(* IEC 61131-3 sources: Lasal-MCP/examples/SampleSource/LASALScreenAdvancedSolution/LASALScreenAdvancedSolution/LASALScreenAdvacnedSolution/Stations/Terminal/HMI/Class/DataRecord, 1 file *)

(* ---- DataRecord.st ---- *)
(*!
<Class
	Name               = "DataRecord"
	Revision           = "0.0"
	RealtimeTask       = "false"
	CyclicTask         = "false"
	BackgroundTask     = "false"
	Sigmatek           = "false"
	OSInterface        = "false"
	HighPriority       = "false"
	Automatic          = "false"
	UpdateMode         = "Prescan"
	SharedCommandTable = "true"
	Objectsize         = "(450,360)">
	<Channels>
		<Server Name="CoordX" Visualized="true" Initialize="false" WriteProtected="true" Retentive="false"/>
		<Server Name="CoordY" Visualized="true" Initialize="false" WriteProtected="true" Retentive="false"/>
		<Server Name="IntError" Visualized="false" Initialize="false" WriteProtected="true" Retentive="false"/>
		<Client Name="_Grafix" Required="false" Internal="false"/>
		<Client Name="_StdLib" Required="false" Internal="false"/>
		<Client Name="AllocateSize" Required="false" Internal="false" DefValue="4 KB"/>
	</Channels>
	<Network Name="DataRecord">
		<!-- List of Components in this network -->
		<Components>
			<Object
				Name       = "_base"
				Class      = "_MyIO"
				Position   = "(218,120)"
				Visualized = "true"
				Remotely   = "true">
				<Channels>
					<Server Name="Refresh"/>
					<Server Name="Server0"/>
					<Client Name="Graphic"/>
					<Client Name="Lse"/>
				</Channels>
			</Object>
		</Components>
		<Comments>
		</Comments>
		<!-- List of Connections in this network -->
		<Connections>
			<Connection Source="this.Server0" Destination="_base.Server0" Vertices="(706,210),(534,210),"/>
			<Connection Source="this.Refresh" Destination="_base.Refresh" Vertices="(706,270),(534,270),"/>
			<Connection Source="_base.Lse" Destination="this.Lse" Vertices="(218,210),(38,210),"/>
		</Connections>
		<!-- Headerfiles -->
		<Options>
		</Options>
	</Network>
</Class>
*)
#pragma using _MyIO

DataRecord : CLASS
: _MyIO
  //Servers:
	CoordX 	: SvrCh_DINT;
	CoordY 	: SvrCh_DINT;
	IntError 	: SvrCh_DINT;
  //Clients:
	_Grafix 	: CltChCmd__Grafix;
	_StdLib 	: CltChCmd__StdLib;
	AllocateSize 	: CltCh_UDINT;
  //Variables:
		pStart 	: ^_DOT;
		pCheck 	: ^_DOT;
		pAct 	: ^_DOT;
		NoOfBufferEntries 	: UDINT;
		MaxNoOfBufferEntries 	: UDINT;
		Delete 	: DINT;
		pError 	: ^void;
  //Functions:

	FUNCTION VIRTUAL GLOBAL Init;
				//! <Function Comment="this method will be called once when the focus will be given to this object" Name="GetFocus"/>
	FUNCTION __CDECL VIRTUAL GLOBAL GetFocus
		VAR_INPUT
			pio 	: ^_IO;			//! <Variable Comment="pointer to _IO information" Name="GetFocus.pio"/>
		END_VAR
		VAR_OUTPUT
			retcode (EAX) 	: _DOIT;			//! <Variable Comment="return _IFAILED if you dont want to get the focus on the other hand _IDLE" Name="GetFocus.retcode"/>
		END_VAR;
				//! <Function Comment="this method is called everytime when the input is active and a event occured" Name="GetEvent"/>
	FUNCTION __CDECL VIRTUAL GLOBAL GetEvent
		VAR_INPUT
			ped 	: ^_EDITOR;			//! <Variable Comment="pointer to _EDITOR information" Name="GetEvent.ped"/>
			pe 	: ^_EVENT;			//! <Variable Comment="pointer to _EVENT information" Name="GetEvent.pe"/>
		END_VAR
		VAR_OUTPUT
			retcode (EAX) 	: _DOIT;			//! <Variable Comment="for the returnstatement there are 3 different possibilities&#13;&#10;  _IDLE ..... the system should goon like it is (system goes on)&#13;&#10;  _IDIDIT ... i did it (system is ready)&#13;&#10;  _IFAILED .. i tried to do my best, but i failed (system is ready)&#13;&#10;" Name="GetEvent.retcode"/>
		END_VAR;
				//! <Function Comment="this method is called everytime when system wants to redraw the io" Name="Draw"/>
	FUNCTION __CDECL VIRTUAL GLOBAL Draw
		VAR_INPUT
			pio 	: ^_IO;			//! <Variable Comment="pointer to _IO information" Name="Draw.pio"/>
			pr 	: ^_RESULT;			//! <Variable Comment="pointer to _RESULT information" Name="Draw.pr"/>
			pv 	: ^_VARIABLE;			//! <Variable Comment="pointer to io _VARIABLE information" Name="Draw.pv"/>
			input 	: BOOL;			//! <Variable Comment="TRUE it&apos;s an input&#13;&#10;FALSE it&apos;s an output" Name="Draw.input"/>
		END_VAR
		VAR_OUTPUT
			retcode (EAX) 	: _DOIT;			//! <Variable Comment="for the returnstatement there are 3 different possibilities&#13;&#10;  _IDLE ..... the system should goon like it is (system goes on)&#13;&#10;  _IDIDIT ... i did it (system is ready)&#13;&#10;  _IFAILED .. i tried to do my best, but i failed (system is re" Name="Draw.retcode"/>
		END_VAR;
				//! <Function Comment="this method is called everytime when system wants to get data for defined io.&#13;&#10;&#13;&#10;pr ........ &#13;&#10;pio ....... pointer to io information&#13;&#10;pv ........ pointer to io variableinformation&#13;&#10;input ..... TRUE it&apos;s an input / FALSE it&apos;s an output&#13;&#10;&#13;&#10;for the returnstatement there are 3 different possibilities&#13;&#10;_IDLE ..... the system should goon like it is (system goes on)&#13;&#10;_IDIDIT ... i did it (system is ready)&#13;&#10;_IFAILED .. i tried to do my best, but i failed (system is ready)&#13;&#10;&#13;&#10;if you want to do it let&apos;s return _IDIDIT and initialize the  structure _RESULT&#13;&#10;" Name="GetData"/>
	FUNCTION __CDECL VIRTUAL GLOBAL GetData
		VAR_INPUT
			pr 	: ^_RESULT;			//! <Variable Comment="pointer to _RESULT information" Name="GetData.pr"/>
			pio 	: ^_IO;			//! <Variable Comment="pointer to _IO information" Name="GetData.pio"/>
			pv 	: ^_VARIABLE;			//! <Variable Comment="pointer to _VARIABLE information given by LSE" Name="GetData.pv"/>
			input 	: BOOL;			//! <Variable Comment="TRUE it&apos;s an input&#13;&#10;FALSE it&apos;s an output" Name="GetData.input"/>
		END_VAR
		VAR_OUTPUT
			retcode (EAX) 	: _DOIT;			//! <Variable Comment="for the returnstatement there are 3 different possibilities&#13;&#10;  _IDLE ..... the system should goon like it is (system goes on)&#13;&#10;  _IDIDIT ... i did it (system is ready)&#13;&#10;  _IFAILED .. i tried to do my best, but i failed (system is ready)" Name="GetData.retcode"/>
		END_VAR;
  //Tables:
	FUNCTION @STD
		VAR_OUTPUT
			ret_code	: CONFSTATES;
		END_VAR;
	FUNCTION GLOBAL TAB @CT_;
END_CLASS;

#pragma usingLtd _Grafix
#pragma usingLtd _StdLib

FUNCTION VIRTUAL GLOBAL DataRecord::Init

  if _FirstScan then

    MaxNoOfBufferEntries := AllocateSize / sizeof(_DOT);

    pStart$^void := _StdLib.MallocV1(size0:= AllocateSize,
                                     mark0:= 0);

    if (pStart = NIL) then
      IntError := -1;
      return;
    else

      pError := _StdLib.MemSet(dest:= pStart,
                               value:= 0,
                               size:= AllocateSize);

      if (pError <> pStart) then
        IntError := -2;
        return;
      end_if;

    end_if;

    Delete := TRUE;
  end_if;

END_FUNCTION

FUNCTION __CDECL VIRTUAL GLOBAL DataRecord::GetEvent
	VAR_INPUT
		ped 	: ^_EDITOR;
		pe 	: ^_EVENT;
	END_VAR
	VAR_OUTPUT
		retcode (EAX) 	: _DOIT;
	END_VAR

  _MyIO::GetEvent(ped:=ped, pe:=pe);

  retcode := _IDLE;

  if (pe^.ftype = _EVENT_HIDMOVE) then

    Delete := FALSE;

    if ((pe^.dot.x > ped^.input.io.space.xy1.x) &
        (pe^.dot.x < ped^.input.io.space.xy2.x) &
        (pe^.dot.y > ped^.input.io.space.xy1.y) &
        (pe^.dot.y < ped^.input.io.space.xy2.y)) then

        retcode := _IDIDIT;

        CoordX := pe^.dot.x - ped^.input.io.space.xy1.x;
        CoordY := pe^.dot.y - ped^.input.io.space.xy1.y;

        if (NoOfBufferEntries >= MaxNoOfBufferEntries) then
          NoOfBufferEntries := 0;

          pAct := pStart;
        end_if;

        pAct^.x := pe^.dot.x;
        pAct^.y := pe^.dot.y;

        pAct := pAct + sizeof(_DOT);
        NoOfBufferEntries += 1;
     end_if;

  elsif (pe^.ftype = _EVENT_HIDRELEASE) then
    Delete := TRUE;
  end_if;

END_FUNCTION

FUNCTION __CDECL VIRTUAL GLOBAL DataRecord::Draw
	VAR_INPUT
		pio 	: ^_IO;
		pr 	: ^_RESULT;
		pv 	: ^_VARIABLE;
		input 	: BOOL;
	END_VAR
	VAR_OUTPUT
		retcode (EAX) 	: _DOIT;
	END_VAR
  VAR
  	act : _NEWSCREEN;
    pNext : ^_DOT;
    bgColor, recordColor : _COLOR;
  END_VAR

  _MyIO::Draw(pio:=pio, pr:=pr, pv:=pv, input:=input);

  push_screen(p0:=#act);

  if (Delete = TRUE) then

    bgColor := _Grafix.MakeColor(backcolor:= pio^.colback,
                                 frontcolor:= pio^.colback);

    _Grafix.Beam(x0:= pio^.space.xy1.x,
                 y0:= pio^.space.xy1.y,
                 x1:= pio^.space.xy2.x,
                 y1:= pio^.space.xy2.y,
                 attrib:= pio^.attrib,
                 color:= bgColor);

  end_if;

  if (pAct <> NIL) then
    pCheck := pStart;
    while (pCheck < (pAct - sizeof(_DOT))) do

      pNext := pCheck + sizeof(_DOT);

      recordColor := _Grafix.MakeColor(backcolor:= pio^.coltxt,
                                       frontcolor:= pio^.coltxt);

      _Grafix.Line(x0:= pCheck^.x,
                   y0:= pCheck^.y,
                   x1:= pNext^.x,
                   y1:= pNext^.y,
                   attrib:= pio^.attrib,
                   color:= recordColor);

      pCheck += sizeof(_DOT);

    end_while;

  end_if;

  pop_screen(p0:=#act);
  copy_screen(p0:=#act, p1:=#pio^.space);

  retcode := _IDIDIT;

END_FUNCTION

FUNCTION __CDECL VIRTUAL GLOBAL DataRecord::GetFocus
	VAR_INPUT
		pio 	: ^_IO;
	END_VAR
	VAR_OUTPUT
		retcode (EAX) 	: _DOIT;
	END_VAR

  _MyIO::GetFocus(pio:=pio);

  pAct := pStart;
  pCheck  := pStart;
  NoOfBufferEntries := 0;

  retcode := _IDLE;

END_FUNCTION

FUNCTION __CDECL VIRTUAL GLOBAL DataRecord::GetData
	VAR_INPUT
		pr 	: ^_RESULT;
		pio 	: ^_IO;
		pv 	: ^_VARIABLE;
		input 	: BOOL;
	END_VAR
	VAR_OUTPUT
		retcode (EAX) 	: _DOIT;
	END_VAR

  _MyIO::GetData(pr:=pr, pio:=pio, pv:=pv, input:=input);

  pr^.value := to_dint((to_udint(CoordX)rol 1)xor(to_udint(CoordY)));

  retcode := _IDIDIT;

END_FUNCTION
